Fanuc KAREL source: kt00488.KL

-- PROVISIONAL review KL for V770-1; original PC SHA256 f1822f571ad6df383e4c57a6869dad4a85f656b5b17265bbc8cb7fe331af00cc
-- Incomplete behavior may be omitted. Consult companion uncertainty JSON. Do not deploy.
PROGRAM KT00488
%NOLOCKGROUP
VAR
  OUT : BOOLEAN
-- UNRESOLVED_DECL P1 type=000101
-- UNRESOLVED_DECL P2 type=000199
BEGIN
  -- UNRESOLVED_PC offsets 5-33; opcodes 49,49,7E,AC,23
  -- UNRESOLVED_PC offsets 38-42; opcodes 7F
END KT00488
